(* Logix 5000 project; controller TFF vendor 1 type 14 code 107 rev 34.11; software revision 34.03; part 15 of 36 *)
(* tags used below, declared in another part *)
   AutoRunTimer : TIMER;   // Auto Run Timer
   Clear : BOOL;   // Clear Operation Table Flag
   DownloadONS : BOOL;
   ErrorCheck : BOOL;   // Error Check Flag
   PhaseClear : BOOL;   // Phase Clear
   PreRunLog : BOOL;   // Log Pre Run Set Points
   ResumeDownloadFromHOLD : BOOL;
   Run : BOOL;   // Operation Run Status
   RunONS : BOOL;   // Run Command One-Shot
   Structure : DINT;   // Structure code
   Value : REAL;   // Temp Value
   AlarmControl : AlarmControl;   // Alarm Control
   AnalogPoint : AnalogInput[50];   // Analog Input Array
   CCPSystem : CCPSystem;   // CCP System Data
   CPU_Scanning : BOOL;   // System Scanning Flag
   Memory_Data : Memory_Data;
   Memory_Message : MESSAGE;   // Data for Message instruction read Memory informations
   Memory_Temp : INT[29];   // Destination elements for message read Memory informations
   MiscREAL : REAL[50];   // Misc Real Values
   Operation : Operation[6,251];   // Operation Table
   PCDateTime : DINT[7];   // Date/Time Array from PC
   Phase : Phases[6];   // Phase Control Array
   Phase0 : ALIAS FOR Phase[0];   // Phase 0
   PhaseTotalizer : PhaseTotalizer[18];   // Phase Totalizers Array
   PLCFault : FaultRecordType;   // PLC Major Fault Record
   Prompt0 : ALIAS FOR Prompt[0];   // Phase 0 Prompt
   Prompt1 : ALIAS FOR Prompt[1];   // Phase 1 Prompt
   Prompt2 : ALIAS FOR Prompt[2];   // Phase 2 Prompt
   Prompt3 : ALIAS FOR Prompt[3];   // Phase 3 Prompt
   Prompt4 : ALIAS FOR Prompt[4];   // Phase 4 Prompt
   Prompt5 : ALIAS FOR Prompt[5];   // Phase 5 Prompt
   TimerControl : TimerControl;   // Timer Control
   Timers : Timers[22];   // Timer Array
   Totalizer : Totalizers[20];   // Totalizers Array
   YA10 : ALIAS FOR DigitalPoint[59];   // PLC Program Major Fault
(* CCPSystem, continued *)

ROUTINE Start   (* ladder *)
// Operation Start Routine
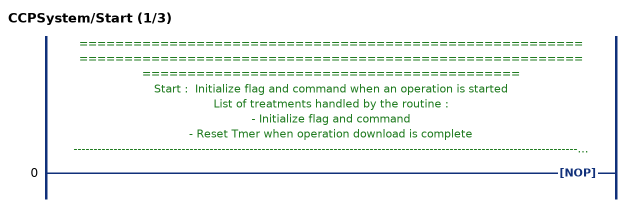
   // ==========================================================================================================================================================
   //                                                                                                      Start :  Initialize flag and command when an operation is started
   //                                                     List of treatments handled by the routine :
   //                                                          - Initialize flag and command
   //                                                          - Reset Tmer when operation download is complete
   //                                                     -----------------------------------------------------------------------------------------------------------------------------------------------------
   //                                                     History
   //                                                         2019-AUG-13 - Actemium - B. Roch - Initial version for Candidate Release 3.00.00.00.a
   // ========================================================================================================================================================
   0: NOP();
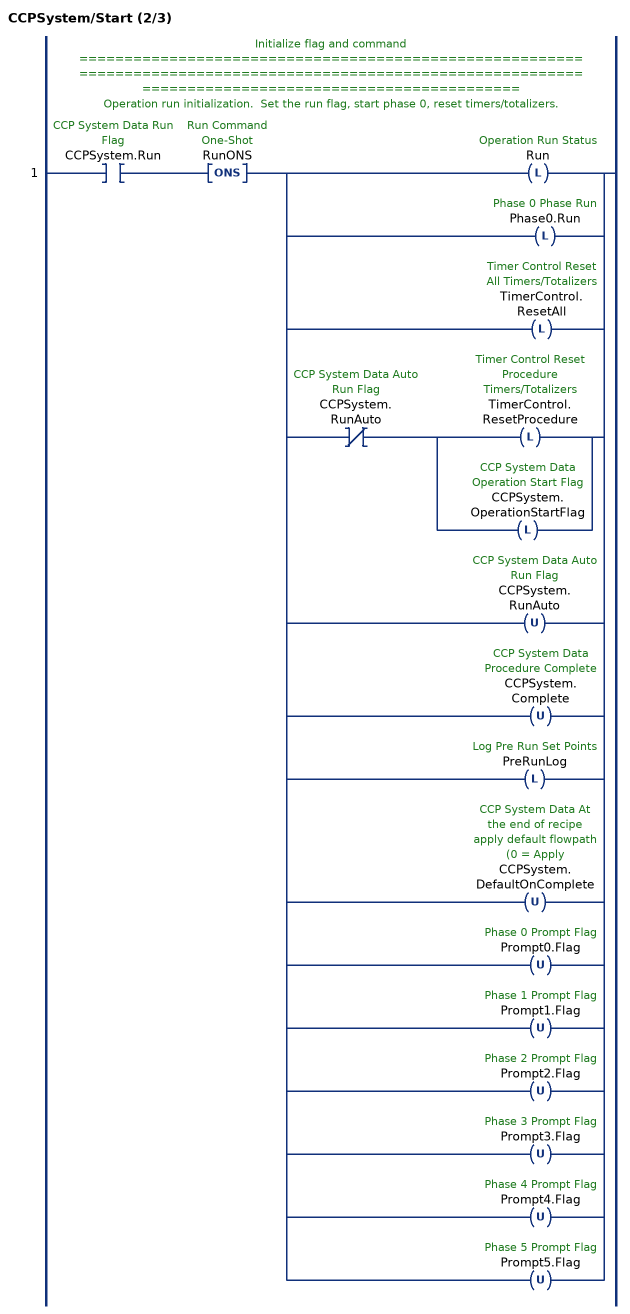
   // Initialize flag and command
   // ==========================================================================================================================================================
   // Operation run initialization.  Set the run flag, start phase 0, reset timers/totalizers.
   1: XIC(CCPSystem.Run)ONS(RunONS)[OTL(Run) ,OTL(Phase0.Run) ,OTL(TimerControl.ResetAll) ,XIO(CCPSystem.RunAuto) [OTL(TimerControl.ResetProcedure) ,OTL(CCPSystem.OperationStartFlag) ] ,OTU(CCPSystem.RunAuto) ,OTU(CCPSystem.Complete) ,OTL(PreRunLog) ,OTU(CCPSystem.DefaultOnComplete) ,OTU(Prompt0.Flag) ,OTU(Prompt1.Flag) ,OTU(Prompt2.Flag) ,OTU(Prompt3.Flag) ,OTU(Prompt4.Flag) ,OTU(Prompt5.Flag) ];
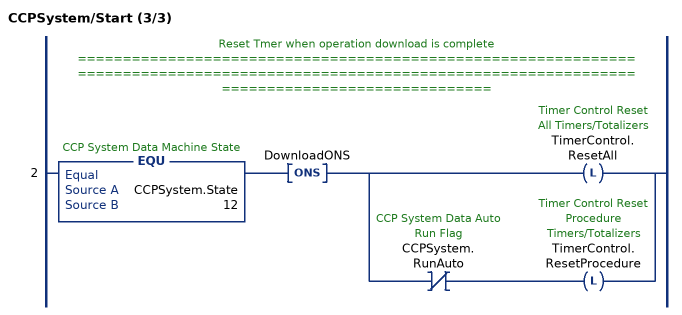
   // Reset Tmer when operation download is complete
   // ==========================================================================================================================================================
   2: EQU(CCPSystem.State,12)ONS(DownloadONS)[OTL(TimerControl.ResetAll) ,XIO(CCPSystem.RunAuto) OTL(TimerControl.ResetProcedure) ];
END_ROUTINE

ROUTINE State   (* ladder *)
// Machine State Routine
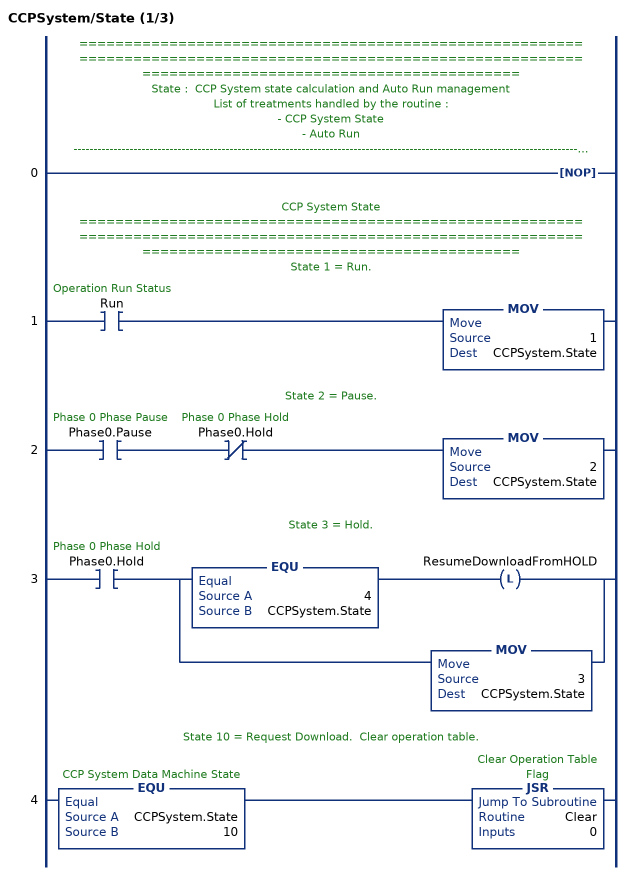
   // ==========================================================================================================================================================
   //                                                                                                  State :  CCP System state calculation and Auto Run management
   //                                                     List of treatments handled by the routine :
   //                                                          - CCP System State
   //                                                          - Auto Run
   //                                                     -----------------------------------------------------------------------------------------------------------------------------------------------------
   //                                                     History
   //                                                         2019-AUG-13 - Actemium - B. Roch - Initial version for Candidate Release 3.00.00.00.a
   //                                       2020-NOV-24 - Merck - Q.SPINDLER - Modifications for Candidate Release 3.00.00.01.b
   //                                     - Restore the State to 4 after hold when it was 4 and hold happen
   // ========================================================================================================================================================
   0: NOP();
   // CCP System State
   // ==========================================================================================================================================================
   // State 1 = Run.
   1: XIC(Run)MOV(1,CCPSystem.State);
   // State 2 = Pause.
   2: XIC(Phase0.Pause)XIO(Phase0.Hold)MOV(2,CCPSystem.State);
   // State 3 = Hold.
   3: XIC(Phase0.Hold)[EQU(4,CCPSystem.State) OTL(ResumeDownloadFromHOLD) ,MOV(3,CCPSystem.State) ];
   // State 10 = Request Download.  Clear operation table.
   4: EQU(CCPSystem.State,10)JSR(Clear,0);
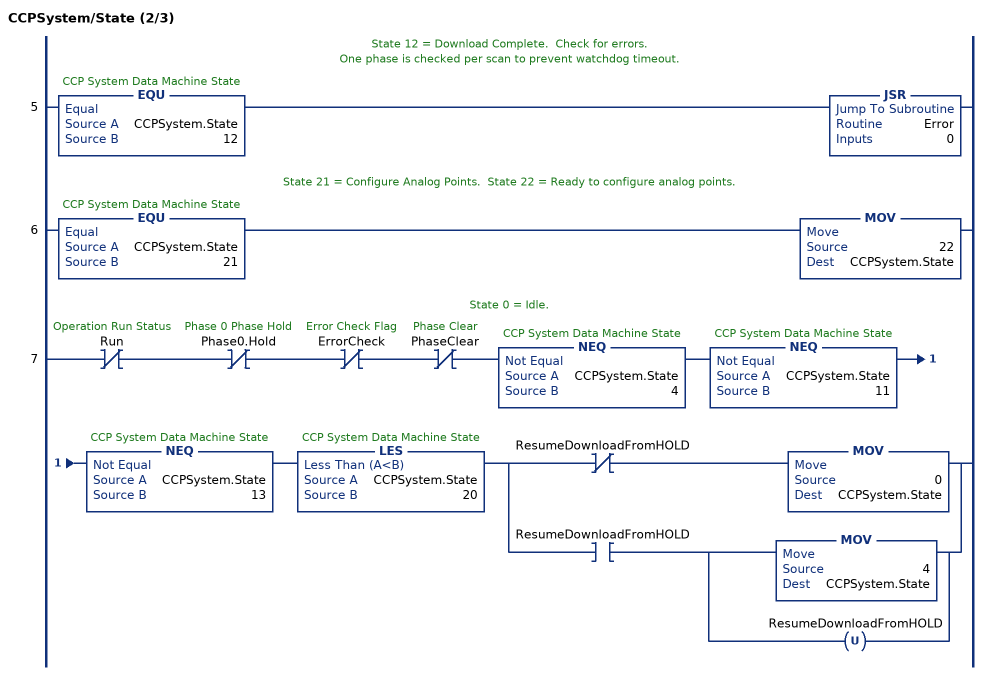
   // State 12 = Download Complete.  Check for errors.
   // One phase is checked per scan to prevent watchdog timeout.
   5: EQU(CCPSystem.State,12)JSR(Error,0);
   // State 21 = Configure Analog Points.  State 22 = Ready to configure analog points.
   6: EQU(CCPSystem.State,21)MOV(22,CCPSystem.State);
   // State 0 = Idle.
   7: XIO(Run)XIO(Phase0.Hold)XIO(ErrorCheck)XIO(PhaseClear)NEQ(CCPSystem.State,4)NEQ(CCPSystem.State,11)NEQ(CCPSystem.State,13)LES(CCPSystem.State,20)[XIO(ResumeDownloadFromHOLD) MOV(0,CCPSystem.State) ,XIC(ResumeDownloadFromHOLD) [MOV(4,CCPSystem.State) ,OTU(ResumeDownloadFromHOLD) ] ];
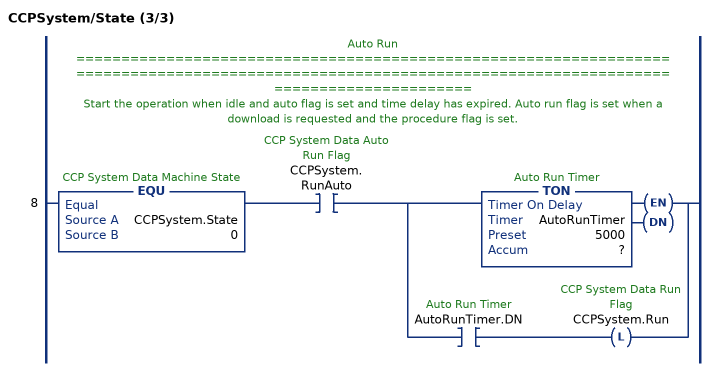
   // Auto Run
   // ==========================================================================================================================================================
   // Start the operation when idle and auto flag is set and time delay has expired. Auto run flag is set when a download is requested and the procedure flag is set.
   8: EQU(CCPSystem.State,0)XIC(CCPSystem.RunAuto)[TON(AutoRunTimer,?,?) ,XIC(AutoRunTimer.DN) OTL(CCPSystem.Run) ];
END_ROUTINE
END_PROGRAM

PROGRAM ControllerFaultRoutine   (* main routine FaultRoutine *)

ROUTINE FaultRoutine   (* ladder *)
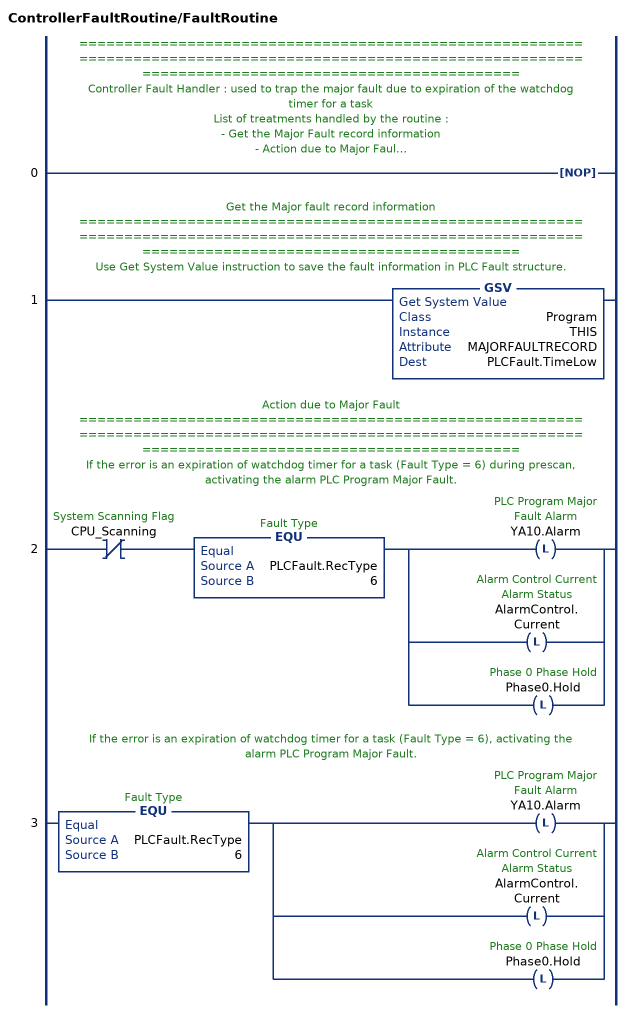
   // ==========================================================================================================================================================
   //                                                                                 Controller Fault Handler : used to trap the major fault due to expiration of the watchdog timer for a task
   //                                                     List of treatments handled by the routine :
   //                                                          - Get the Major Fault record information
   //                                                          - Action due to Major Fault
   //                                                     -----------------------------------------------------------------------------------------------------------------------------------------------------
   //                                                     History
   //                                                          2019-AUG-13 - Actemium - B. Roch - Initial version for Candidate Release 3.00.00.00.a
   // ==========================================================================================================================================================
   0: NOP();
   // Get the Major fault record information
   // ==========================================================================================================================================================
   // Use Get System Value instruction to save the fault information in PLC Fault structure.
   1: GSV(Program,THIS,MAJORFAULTRECORD,PLCFault.TimeLow);
   // Action due to Major Fault
   // ==========================================================================================================================================================
   // If the error is an expiration of watchdog timer for a task (Fault Type = 6) during prescan, activating the alarm PLC Program Major Fault.
   2: XIO(CPU_Scanning)EQU(PLCFault.RecType,6)[OTL(YA10.Alarm) ,OTL(AlarmControl.Current) ,OTL(Phase0.Hold) ];
   // If the error is an expiration of watchdog timer for a task (Fault Type = 6), activating the alarm PLC Program Major Fault.
   3: EQU(PLCFault.RecType,6)[OTL(YA10.Alarm) ,OTL(AlarmControl.Current) ,OTL(Phase0.Hold) ];
END_ROUTINE
END_PROGRAM

PROGRAM MainProgram   (* main routine MainRoutine, fault routine FaultRoutine *)
// Date/Time Synchronization
VAR
   Address : DINT := 9;   // Temp Address used in Time Loop
   AddressTotalizer : DINT := 2;   // Temp Address used in modPhaseTotal
   Index : DINT := 4;   // Index
   PLCDST : SINT;   // Current PLC Day Light Saving
   PLCTimeZoneString : STRING := 'UTC+00:00 Coordinated Universal Time';   // Current PLC TimeZone
   SCL : SCALE := (In := -4.0, InRawMax := 99999.0, InEUMax := 999.99, Out := -0.04, MinAlarm := 1);
   TimeZoneUTC0 : STRING := 'UTC+00:00 Coordinated Universal Time';   // String value for Time zone UTC 0
END_VAR

ROUTINE FaultRoutine   (* ladder *)
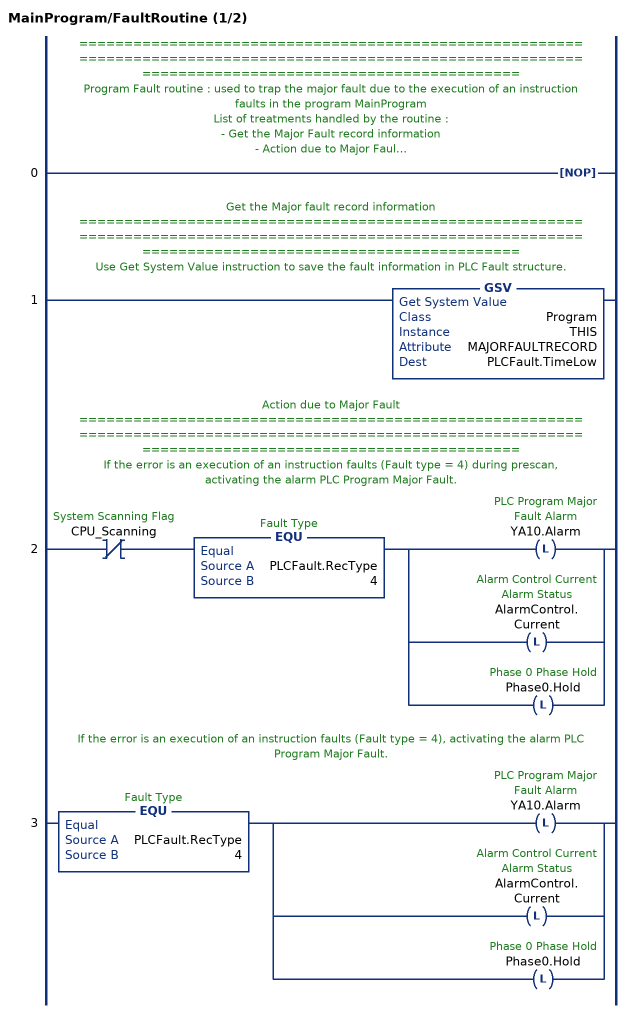
   // ==========================================================================================================================================================
   //                                                               Program Fault routine : used to trap the major fault due to the execution of an instruction faults in the program MainProgram
   //                                                     List of treatments handled by the routine :
   //                                                          - Get the Major Fault record information
   //                                                          - Action due to Major Fault
   //                                                     -----------------------------------------------------------------------------------------------------------------------------------------------------
   //                                                     History
   //                                                         2019-AUG-13 - Actemium - B. Roch - Initial version for Candidate Release 3.00.00.00.a
   // ==========================================================================================================================================================
   0: NOP();
   // Get the Major fault record information
   // ==========================================================================================================================================================
   // Use Get System Value instruction to save the fault information in PLC Fault structure.
   1: GSV(Program,THIS,MAJORFAULTRECORD,PLCFault.TimeLow);
   // Action due to Major Fault
   // ==========================================================================================================================================================
   // If the error is an execution of an instruction faults (Fault type = 4) during prescan, activating the alarm PLC Program Major Fault.
   2: XIO(CPU_Scanning)EQU(PLCFault.RecType,4)[OTL(YA10.Alarm) ,OTL(AlarmControl.Current) ,OTL(Phase0.Hold) ];
   // If the error is an execution of an instruction faults (Fault type = 4), activating the alarm PLC Program Major Fault.
   3: EQU(PLCFault.RecType,4)[OTL(YA10.Alarm) ,OTL(AlarmControl.Current) ,OTL(Phase0.Hold) ];
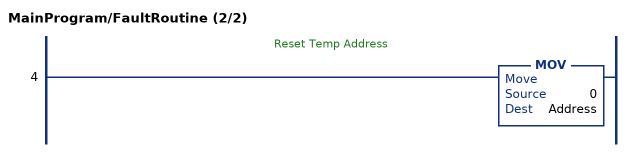
   // Reset Temp Address
   4: MOV(0,Address);
END_ROUTINE

ROUTINE MainRoutine   (* ladder *)
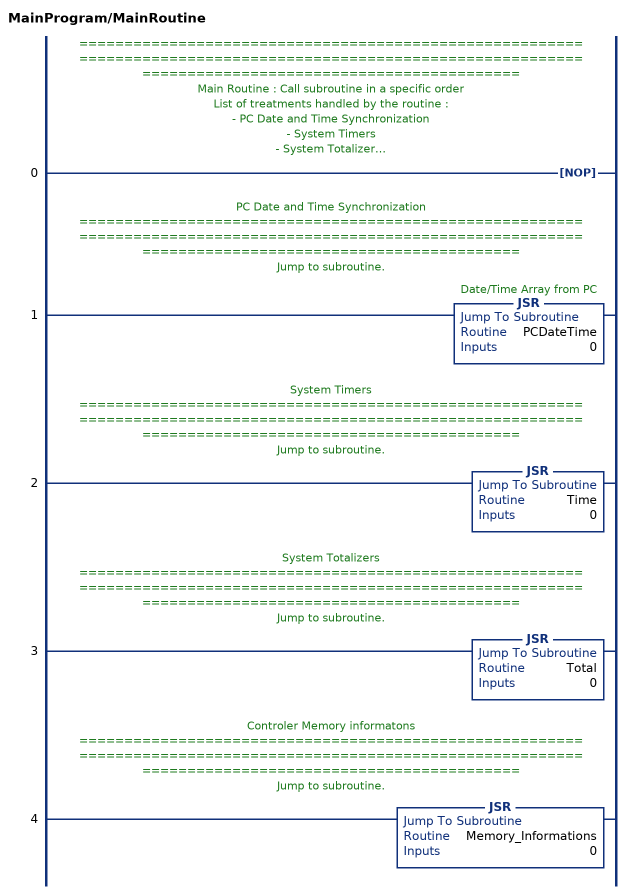
   // ==========================================================================================================================================================
   //                                                                                                            Main Routine : Call subroutine in a specific order
   //                                                     List of treatments handled by the routine :
   //                                                          - PC Date and Time Synchronization
   //                                                          - System Timers
   //                                                          - System Totalizers
   //                                                           - Controler Memory informatons
   //                                                     -----------------------------------------------------------------------------------------------------------------------------------------------------
   //                                                     History
   //                                                       2019-AUG-13 - Actemium - B. Roch - Initial version for Candidate Release 3.00.00.00.a
   //                                                        2020-SEP-24 - Merck - Q. Spindler - Modifications for Candidate Release 3.00.00.01.a
   // 			- Add Memory_Information routine call
   // ==========================================================================================================================================================
   0: NOP();
   // PC Date and Time Synchronization
   // ==========================================================================================================================================================
   // Jump to subroutine.
   1: JSR(PCDateTime,0);
   // System Timers
   // ==========================================================================================================================================================
   // Jump to subroutine.
   2: JSR(Time,0);
   // System Totalizers
   // ==========================================================================================================================================================
   // Jump to subroutine.
   3: JSR(Total,0);
   // Controler Memory informatons
   // ==========================================================================================================================================================
   // Jump to subroutine.
   4: JSR(Memory_Informations,0);
END_ROUTINE

ROUTINE Memory_Data   (* ladder *)
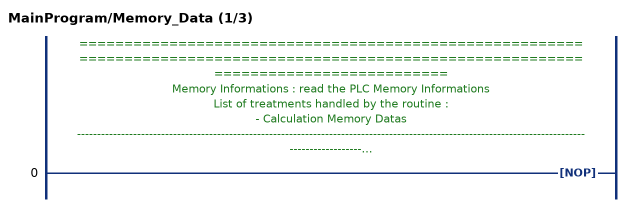
   // ==========================================================================================================================================
   // Memory Informations : read the PLC Memory Informations
   // List of treatments handled by the routine :
   // - Calculation Memory Datas
   //                                                     --------------------------------------------------------------------------------------------------------------------------------------------------
   // History
   // 		2020-SEP-24 - Merck - Q. Spindler - Initial version for Candidate Release 3.00.00.01.a
   // ==========================================================================================================================================
   0: NOP();
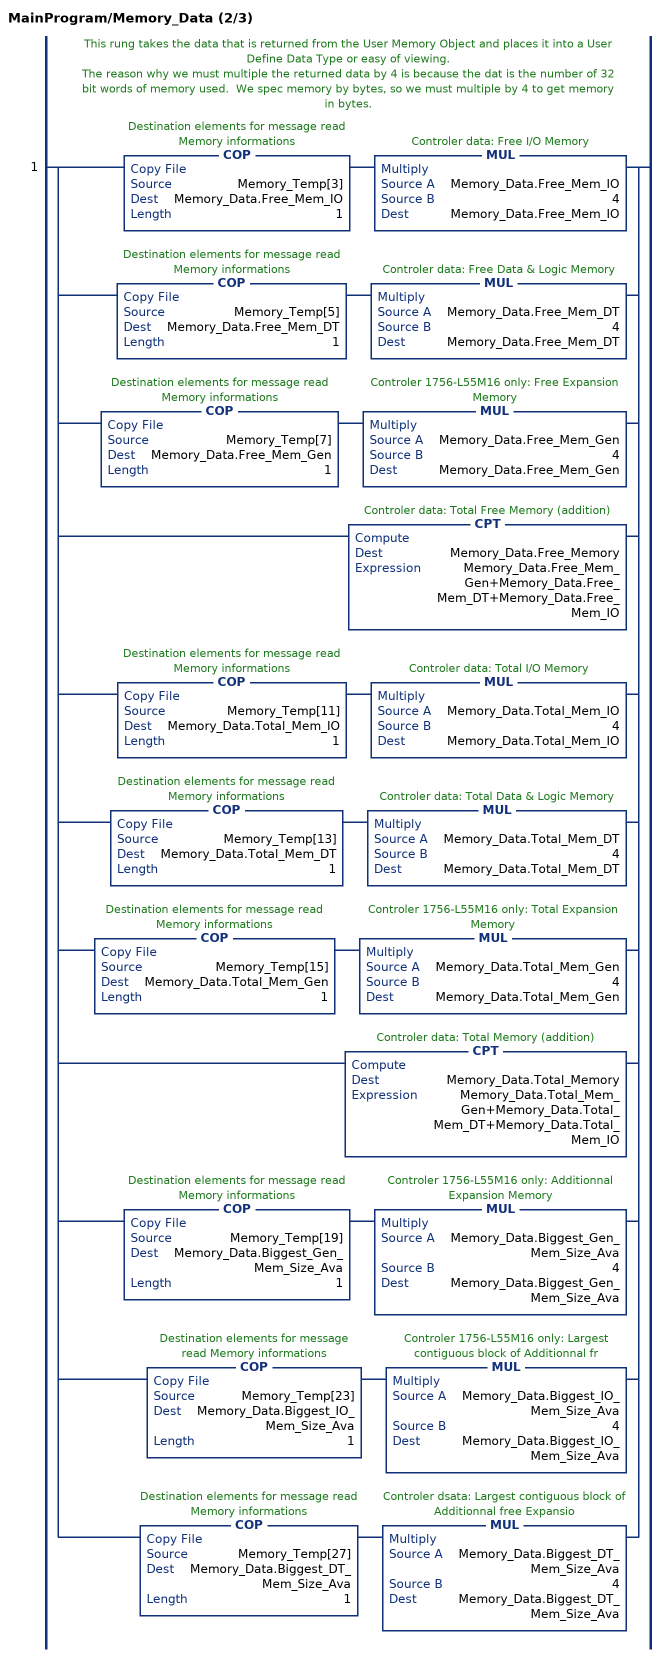
   // This rung takes the data that is returned from the User Memory Object and places it into a User Define Data Type or easy of viewing.
   // The reason why we must multiple the returned data by 4 is because the dat is the number of 32 bit words of memory used.  We spec memory by bytes, so we must multiple by 4 to get memory in bytes.
   1: [COP(Memory_Temp[3],Memory_Data.Free_Mem_IO,1) MUL(Memory_Data.Free_Mem_IO,4,Memory_Data.Free_Mem_IO) ,COP(Memory_Temp[5],Memory_Data.Free_Mem_DT,1) MUL(Memory_Data.Free_Mem_DT,4,Memory_Data.Free_Mem_DT) ,COP(Memory_Temp[7],Memory_Data.Free_Mem_Gen,1) MUL(Memory_Data.Free_Mem_Gen,4,Memory_Data.Free_Mem_Gen) ,CPT(Memory_Data.Free_Memory,Memory_Data.Free_Mem_Gen+Memory_Data.Free_Mem_DT+Memory_Data.Free_Mem_IO) ,COP(Memory_Temp[11],Memory_Data.Total_Mem_IO,1) MUL(Memory_Data.Total_Mem_IO,4,Memory_Data.Total_Mem_IO) ,COP(Memory_Temp[13],Memory_Data.Total_Mem_DT,1) MUL(Memory_Data.Total_Mem_DT,4,Memory_Data.Total_Mem_DT) ,COP(Memory_Temp[15],Memory_Data.Total_Mem_Gen,1) MUL(Memory_Data.Total_Mem_Gen,4,Memory_Data.Total_Mem_Gen) ,CPT(Memory_Data.Total_Memory,Memory_Data.Total_Mem_Gen+Memory_Data.Total_Mem_DT+Memory_Data.Total_Mem_IO) ,COP(Memory_Temp[19],Memory_Data.Biggest_Gen_Mem_Size_Ava,1) MUL(Memory_Data.Biggest_Gen_Mem_Size_Ava,4,Memory_Data.Biggest_Gen_Mem_Size_Ava) ,COP(Memory_Temp[23],Memory_Data.Biggest_IO_Mem_Size_Ava,1) MUL(Memory_Data.Biggest_IO_Mem_Size_Ava,4,Memory_Data.Biggest_IO_Mem_Size_Ava) ,COP(Memory_Temp[27],Memory_Data.Biggest_DT_Mem_Size_Ava,1) MUL(Memory_Data.Biggest_DT_Mem_Size_Ava,4,Memory_Data.Biggest_DT_Mem_Size_Ava) ];
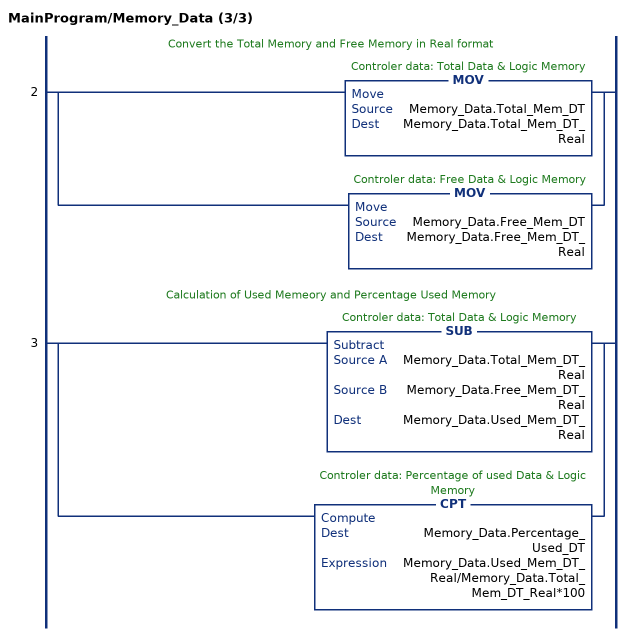
   // Convert the Total Memory and Free Memory in Real format
   2: [MOV(Memory_Data.Total_Mem_DT,Memory_Data.Total_Mem_DT_Real) ,MOV(Memory_Data.Free_Mem_DT,Memory_Data.Free_Mem_DT_Real) ];
   // Calculation of Used Memeory and Percentage Used Memory
   3: [SUB(Memory_Data.Total_Mem_DT_Real,Memory_Data.Free_Mem_DT_Real,Memory_Data.Used_Mem_DT_Real) ,CPT(Memory_Data.Percentage_Used_DT,Memory_Data.Used_Mem_DT_Real/Memory_Data.Total_Mem_DT_Real*100) ];
END_ROUTINE

ROUTINE Memory_Informations   (* ladder *)
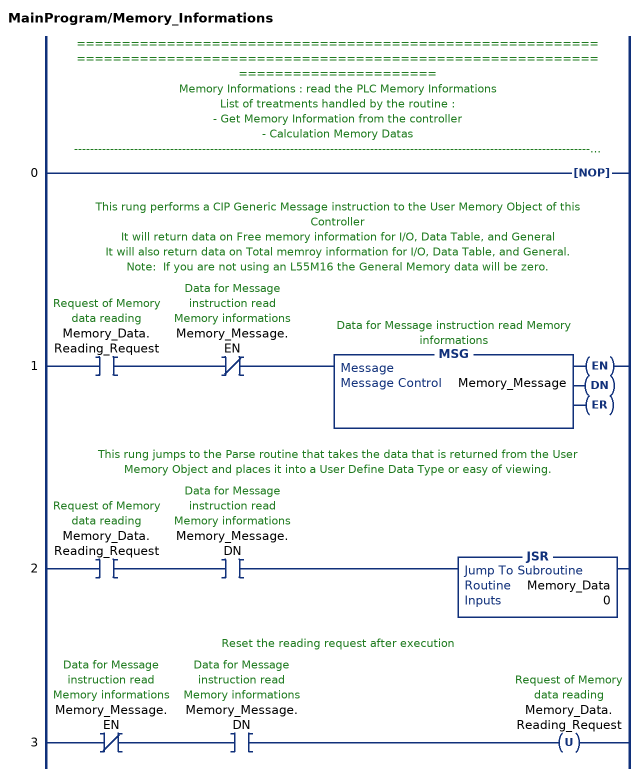
   // ==========================================================================================================================================
   // Memory Informations : read the PLC Memory Informations
   // List of treatments handled by the routine :
   // - Get Memory Information from the controller
   // - Calculation Memory Datas
   //                                                     --------------------------------------------------------------------------------------------------------------------------------------------------
   // History
   // 		2020-SEP-24 - Merck - Q. Spindler - Initial version for Candidate Release 3.00.00.01.a
   // ==========================================================================================================================================
   0: NOP();
   // This rung performs a CIP Generic Message instruction to the User Memory Object of this Controller
   // It will return data on Free memory information for I/O, Data Table, and General
   // It will also return data on Total memroy information for I/O, Data Table, and General.
   // Note:  If you are not using an L55M16 the General Memory data will be zero.
   1: XIC(Memory_Data.Reading_Request)XIO(Memory_Message.EN)MSG(Memory_Message);
   // This rung jumps to the Parse routine that takes the data that is returned from the User Memory Object and places it into a User Define Data Type or easy of viewing.
   2: XIC(Memory_Data.Reading_Request)XIC(Memory_Message.DN)JSR(Memory_Data,0);
   // Reset the reading request after execution
   3: XIO(Memory_Message.EN)XIC(Memory_Message.DN)OTU(Memory_Data.Reading_Request);
END_ROUTINE

ROUTINE modPhaseTotal   (* ladder *)
// Phase Totalizer Module
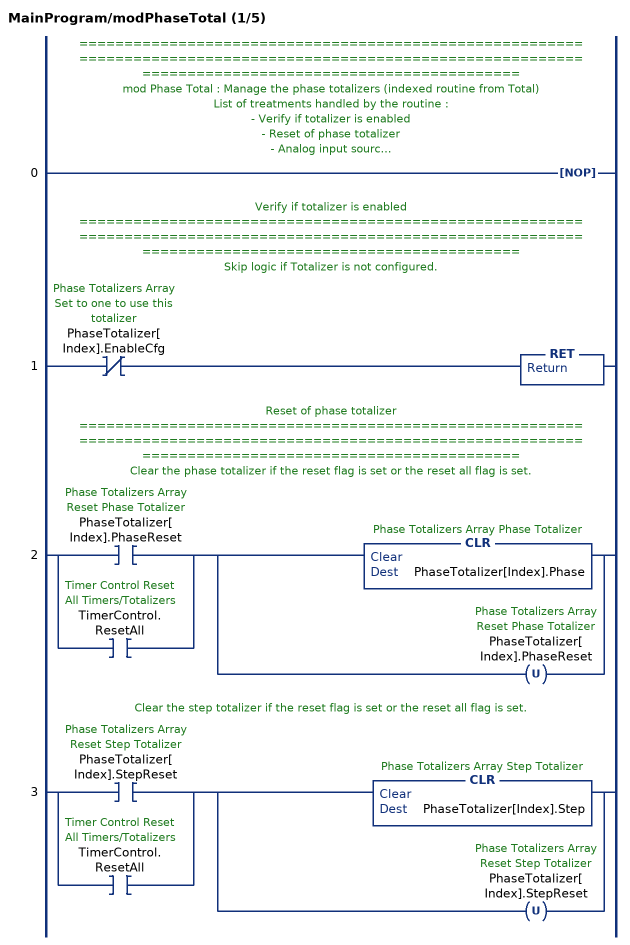
   // ==========================================================================================================================================================
   //                                                                                                   mod Phase Total : Manage the phase totalizers (indexed routine from Total)
   //                                                     List of treatments handled by the routine :
   //                                                          - Verify if totalizer is enabled
   //                                                          - Reset of phase totalizer
   //                                                          - Analog input source
   //                                                          - Calculating the totalizer values
   //                                                     -----------------------------------------------------------------------------------------------------------------------------------------------------
   //                                                     History
   //                                                         2019-AUG-13 - Actemium - B. Roch - Initial version for Candidate Release 3.00.00.00.a
   // ==========================================================================================================================================================
   0: NOP();
   // Verify if totalizer is enabled
   // ==========================================================================================================================================================
   // Skip logic if Totalizer is not configured.
   1: XIO(PhaseTotalizer[Index].EnableCfg)RET();
   // Reset of phase totalizer
   // ==========================================================================================================================================================
   // Clear the phase totalizer if the reset flag is set or the reset all flag is set.
   2: [XIC(PhaseTotalizer[Index].PhaseReset) ,XIC(TimerControl.ResetAll) ][CLR(PhaseTotalizer[Index].Phase) ,OTU(PhaseTotalizer[Index].PhaseReset) ];
   // Clear the step totalizer if the reset flag is set or the reset all flag is set.
   3: [XIC(PhaseTotalizer[Index].StepReset) ,XIC(TimerControl.ResetAll) ][CLR(PhaseTotalizer[Index].Step) ,OTU(PhaseTotalizer[Index].StepReset) ];
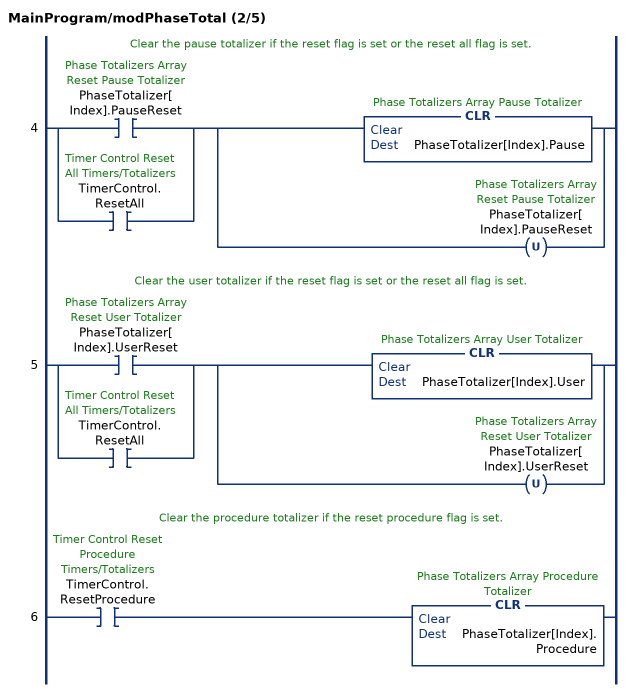
   // Clear the pause totalizer if the reset flag is set or the reset all flag is set.
   4: [XIC(PhaseTotalizer[Index].PauseReset) ,XIC(TimerControl.ResetAll) ][CLR(PhaseTotalizer[Index].Pause) ,OTU(PhaseTotalizer[Index].PauseReset) ];
   // Clear the user totalizer if the reset flag is set or the reset all flag is set.
   5: [XIC(PhaseTotalizer[Index].UserReset) ,XIC(TimerControl.ResetAll) ][CLR(PhaseTotalizer[Index].User) ,OTU(PhaseTotalizer[Index].UserReset) ];
   // Clear the procedure totalizer if the reset procedure flag is set.
   6: XIC(TimerControl.ResetProcedure)CLR(PhaseTotalizer[Index].Procedure);
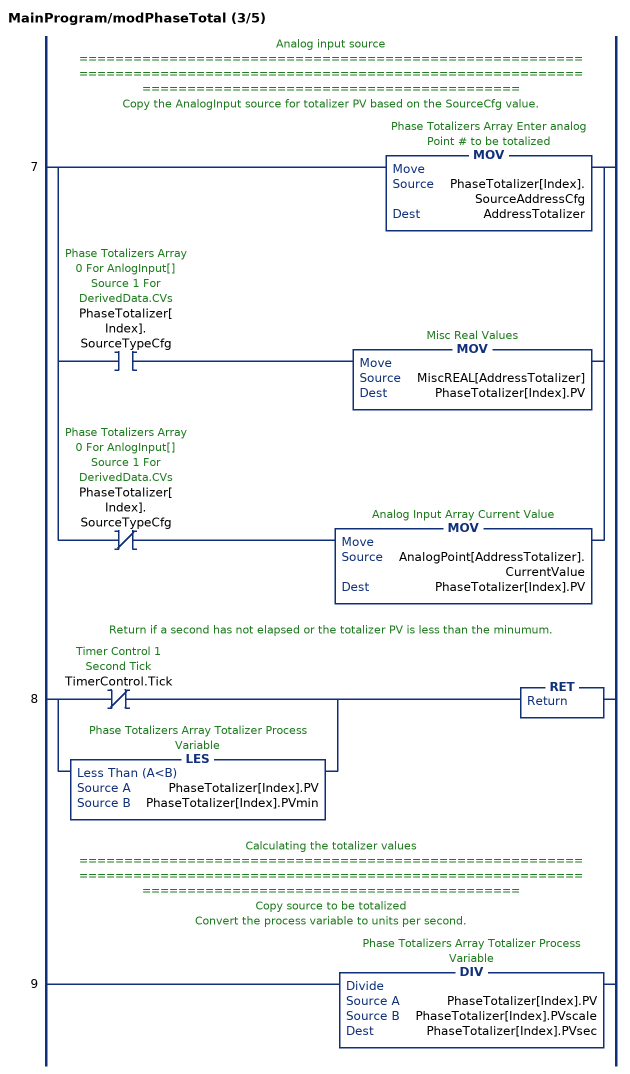
   // Analog input source
   // ==========================================================================================================================================================
   // Copy the AnalogInput source for totalizer PV based on the SourceCfg value.
   7: [MOV(PhaseTotalizer[Index].SourceAddressCfg,AddressTotalizer) ,XIC(PhaseTotalizer[Index].SourceTypeCfg) MOV(MiscREAL[AddressTotalizer],PhaseTotalizer[Index].PV) ,XIO(PhaseTotalizer[Index].SourceTypeCfg) MOV(AnalogPoint[AddressTotalizer].CurrentValue,PhaseTotalizer[Index].PV) ];
   // Return if a second has not elapsed or the totalizer PV is less than the minumum.
   8: [XIO(TimerControl.Tick) ,LES(PhaseTotalizer[Index].PV,PhaseTotalizer[Index].PVmin) ]RET();
   // Calculating the totalizer values
   // ==========================================================================================================================================================
   // Copy source to be totalized
   // Convert the process variable to units per second.
   9: DIV(PhaseTotalizer[Index].PV,PhaseTotalizer[Index].PVscale,PhaseTotalizer[Index].PVsec);
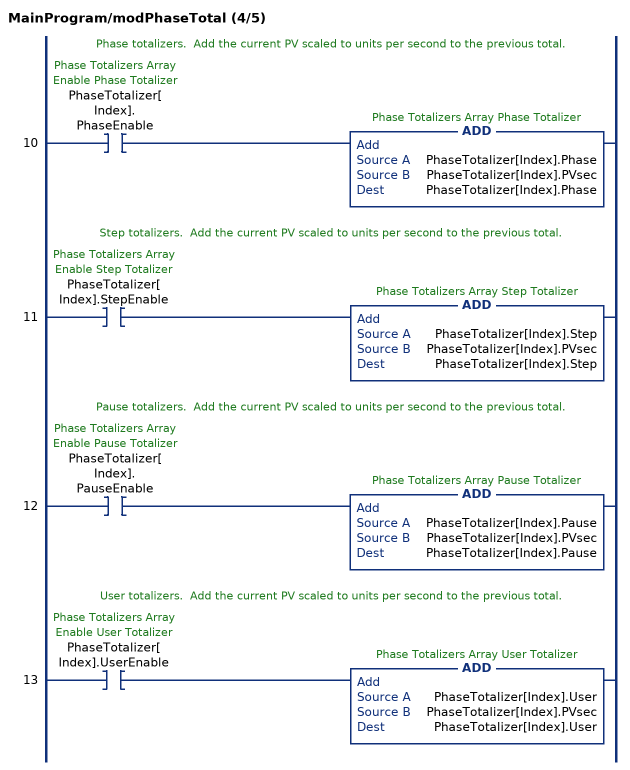
   // Phase totalizers.  Add the current PV scaled to units per second to the previous total.
   10: XIC(PhaseTotalizer[Index].PhaseEnable)ADD(PhaseTotalizer[Index].Phase,PhaseTotalizer[Index].PVsec,PhaseTotalizer[Index].Phase);
   // Step totalizers.  Add the current PV scaled to units per second to the previous total.
   11: XIC(PhaseTotalizer[Index].StepEnable)ADD(PhaseTotalizer[Index].Step,PhaseTotalizer[Index].PVsec,PhaseTotalizer[Index].Step);
   // Pause totalizers.  Add the current PV scaled to units per second to the previous total.
   12: XIC(PhaseTotalizer[Index].PauseEnable)ADD(PhaseTotalizer[Index].Pause,PhaseTotalizer[Index].PVsec,PhaseTotalizer[Index].Pause);
   // User totalizers.  Add the current PV scaled to units per second to the previous total.
   13: XIC(PhaseTotalizer[Index].UserEnable)ADD(PhaseTotalizer[Index].User,PhaseTotalizer[Index].PVsec,PhaseTotalizer[Index].User);
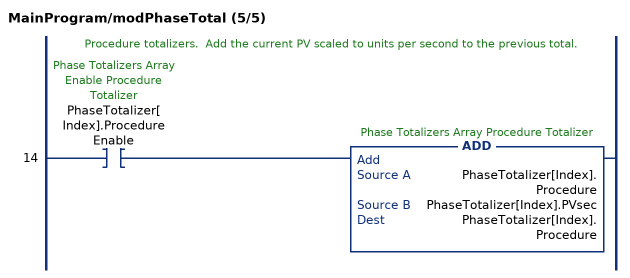
   // Procedure totalizers.  Add the current PV scaled to units per second to the previous total.
   14: XIC(PhaseTotalizer[Index].ProcedureEnable)ADD(PhaseTotalizer[Index].Procedure,PhaseTotalizer[Index].PVsec,PhaseTotalizer[Index].Procedure);
END_ROUTINE
